(* IEC 61131-3 sources: llm-plc-st-eval/data/processed_definitivo/qwen2.5-coder_14b/B8/zero_shot, 3 files *)

(* ---- ejec_1.st ---- *)
FUNCTION_BLOCK FB_Puerta
VAR_INPUT
    puertaAbierta : BOOL; // Entrada que indica si la puerta está abierta
    reset : BOOL; // Entrada para resetear el contador de aperturas
END_VAR

VAR_OUTPUT
    aviso : BOOL; // Salida que indica si se han acumulado 5 o más aperturas
    nAperturas : INT; // Salida que muestra el número de aperturas
END_VAR

VAR
    puertaAbiertaAnterior : BOOL; // Variable para almacenar el estado anterior de puertaAbierta
END_VAR

// Inicialización de variables
IF reset THEN
    nAperturas := 0;
    aviso := FALSE;
    puertaAbiertaAnterior := FALSE;
END_IF

// Detectar transición de FALSE a TRUE en puertaAbierta
IF NOT puertaAbiertaAnterior AND puertaAbierta THEN
    nAperturas := nAperturas + 1;
END_IF

// Actualizar el estado anterior de puertaAbierta
puertaAbiertaAnterior := puertaAbierta;

// Activar la salida de aviso si se han acumulado 5 o más aperturas
IF nAperturas >= 5 THEN
    aviso := TRUE;
ELSE
    aviso := FALSE;
END_IF
END_FUNCTION_BLOCK

(* ---- ejec_2.st ---- *)
FUNCTION_BLOCK FB_Puerta
VAR_INPUT
    puertaAbierta : BOOL; // Entrada que indica si la puerta está abierta
    reset : BOOL; // Entrada para resetear el contador de aperturas
END_VAR

VAR_OUTPUT
    aviso : BOOL; // Salida que indica si se han acumulado 5 o más aperturas
    nAperturas : INT; // Salida que muestra el número de aperturas
END_VAR

VAR
    puertaAbiertaAnterior : BOOL; // Variable para almacenar el estado anterior de puertaAbierta
END_VAR

// Inicialización de variables
IF NOT puertaAbiertaAnterior THEN
    puertaAbiertaAnterior := puertaAbierta;
END_IF

// Lógica de reset
IF reset THEN
    nAperturas := 0;
    aviso := FALSE;
END_IF

// Contador de aperturas
IF puertaAbierta AND NOT puertaAbiertaAnterior THEN
    nAperturas := nAperturas + 1;
END_IF

// Actualización del estado anterior de puertaAbierta
puertaAbiertaAnterior := puertaAbierta;

// Lógica de aviso
IF nAperturas >= 5 THEN
    aviso := TRUE;
ELSE
    aviso := FALSE;
END_IF
END_FUNCTION_BLOCK

(* ---- ejec_3.st ---- *)
FUNCTION_BLOCK FB_Puerta
VAR_INPUT
    puertaAbierta : BOOL; // Entrada que indica si la puerta está abierta
    reset : BOOL; // Entrada para resetear el contador de aperturas
END_VAR

VAR_OUTPUT
    aviso : BOOL; // Salida que indica si se han acumulado 5 o más aperturas
    nAperturas : INT; // Salida que muestra el número de aperturas
END_VAR

VAR
    puertaAbiertaAnterior : BOOL := FALSE; // Variable para almacenar el estado anterior de la puerta
END_VAR

// Comprueba si se ha reseteado el sistema
IF reset THEN
    nAperturas := 0; // Reinicia el contador de aperturas
    aviso := FALSE; // Desactiva el aviso
ELSE
    // Comprueba si la puerta ha pasado de cerrada a abierta
    IF NOT puertaAbiertaAnterior AND puertaAbierta THEN
        nAperturas := nAperturas + 1; // Incrementa el contador de aperturas
    END_IF

    // Actualiza el estado anterior de la puerta
    puertaAbiertaAnterior := puertaAbierta;

    // Comprueba si se han acumulado 5 o más aperturas
    IF nAperturas >= 5 THEN
        aviso := TRUE; // Activa el aviso
    ELSE
        aviso := FALSE; // Desactiva el aviso
    END_IF
END_IF
END_FUNCTION_BLOCK
